(*
SPDX-FileCopyrightText: © 2026 Oleksandr Tiutyk <trofimich@gmail.com>
SPDX-License-Identifier: MIT
License: https://opensource.org/license/mit
*)

(*
Reads a fixed-capacity list whose entries borrow live PLC values.

Edit _SourceValue in Watch. The list stores one descriptor for that variable and _Value follows subsequent edits.
The persistent source must outlive the list's use of the entry. No payload ownership is transferred.
Map this program to one dedicated cyclic task. The program performs cleanup for that task.
*)

{attribute 'no_explicit_call' := 'do not call this function block directly'}
PROGRAM BorrowedListExample
VAR
	{attribute 'hide'}
	_ClassName : STRING := __POUNAME();
	_List : TOF_Collections.List<3>(valueValidator := 0);
	_SourceValue : INT := 42;
	_Value : INT;
END_VAR

IF _List.Empty THEN
	_List.AppendGeneric(value := TOF_Core.GenericValueFactory.FromIntReference(value := _SourceValue));
END_IF

_Value := _List.Get(index := 0).AsInt();

TOF_Core.DynamicMemoryManager.RaiseIfAllocationFailed();
TOF_Core.DynamicMemoryManager.CleanupMemory();

// Borrows the initialized program name. Treat it as read-only.
{attribute 'monitoring' := 'call'}
PROPERTY ClassName : REFERENCE TO STRING
GET
ClassName REF= _ClassName;
END_GET
END_PROPERTY

// Borrows the initialized namespace name. Treat it as read-only.
{attribute 'monitoring' := 'call'}
PROPERTY NamespaceName : REFERENCE TO STRING
GET
NamespaceName REF= CurrentNamespace.Name;
END_GET
END_PROPERTY

END_PROGRAM

(* stored: Version 1.1.0.1
   POU BorrowedListExample: Id {e35842cc-8f85-485d-b26c-0f85ad126b3d}, SpecialFunc None
   Property ClassName: Id {7bd129b2-3ed5-42ac-ac8b-5f5ed325e353}
   Get Get: Id {9cef1d48-4e7c-4a91-a336-fd027e4531b6}
   Property NamespaceName: Id {2e4901ec-414a-4385-b751-4b67d97dfbd5}
   Get Get: Id {73293a31-2884-40de-b37d-66ea963eae41} *)
